FUNCTION_BLOCK Status_Remota (* Estado da comunicacao de uma remota Modbus TCP - HidrycoLib *)
  (* Standard: 61499-2 *)
  (* Version 1.1, 06/11/2026, Hidryco, Hidryco, 1.1: Ciclo (E_CYCLE 2 s) pede a leitura do connStatus (Conexao.REQ); estado se corrige sozinho e STS_VIVO vai para a IHM detectar CLP sem dados. 1.0: le o connStatus (online/offline) do escravo MODBUSGENTCPS pelo symlink stsConexao (ligar no hardware: connStatus = RESID.instancia.stsConexao). IThis: STS_ESTADO (0 aguardando, 1 comunicando, 2 sem comunicacao) e STS_COMUNICANDO. *)
  PACKAGE Hidryco.HidrycoLib;
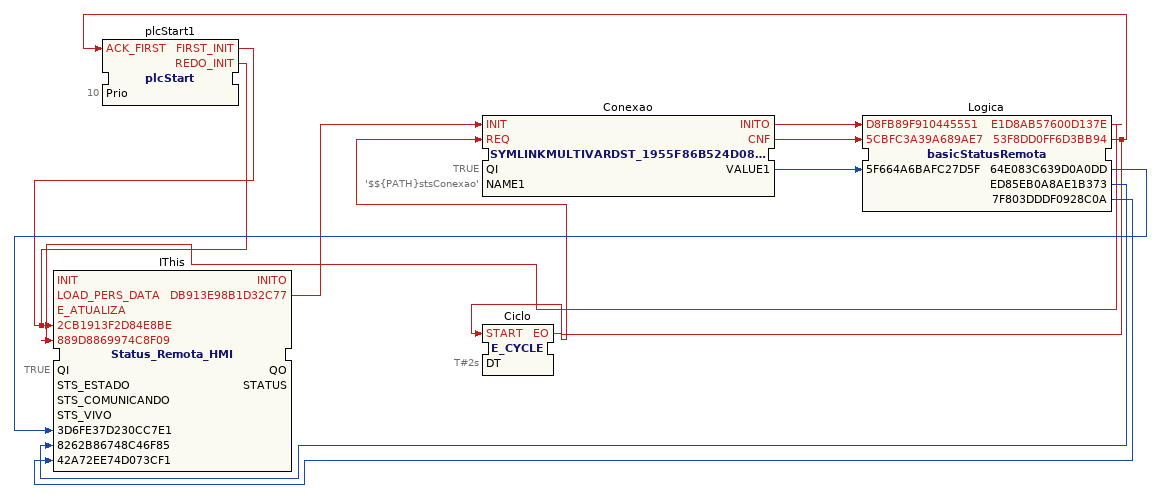
  FBS
    IThis : Status_Remota_HMI(QI := TRUE);
    plcStart1 : plcStart(Prio := 10);
    Conexao : SYMLINKMULTIVARDST_1955F86B524D08A33(QI := TRUE, NAME1 := '$${PATH}stsConexao'); {SET_ATTRIBUTE(Configuration.GenericFBType.InterfaceParams, Runtime.System#I:=1;VALUE${I$}:STRING)}
    Logica : basicStatusRemota;
    Ciclo : E_CYCLE(DT := T#2s);
  END_FBS
  EVENT_CONNECTIONS
    plcStart1.FIRST_INIT TO IThis.2CB1913F2D84E8BE;
    plcStart1.REDO_INIT TO IThis.2CB1913F2D84E8BE;
    IThis.DB913E98B1D32C77 TO Conexao.INIT;
    Conexao.INITO TO Logica.D8FB89F910445551;
    Conexao.CNF TO Logica.5CBFC3A39A689AE7;
    Logica.E1D8AB57600D137E TO IThis.889D8869974C8F09;
    Logica.53F8DD0FF6D3BB94 TO plcStart1.ACK_FIRST;
    Logica.53F8DD0FF6D3BB94 TO Ciclo.START;
    Ciclo.EO TO Conexao.REQ;
  END_CONNECTIONS
  DATA_CONNECTIONS
    Conexao.VALUE1 TO Logica.5F664A6BAFC27D5F;
    Logica.64E083C639D0A0DD TO IThis.3D6FE37D230CC7E1;
    Logica.ED85EB0A8AE1B373 TO IThis.8262B86748C46F85;
    Logica.7F803DDDF0928C0A TO IThis.42A72EE74D073CF1;
  END_CONNECTIONS
END_FUNCTION_BLOCK
